// TIA Portal V20 export
// export: Created 2026-10-20T12:44:30.4346877Z, ExportSetting WithDefaults, DisplayName Totally Integrated Automation Portal, DisplayVersion V20 Update 6, DisplayName TIA Portal Openness, DisplayVersion V20 Update 6, DisplayName TIA Portal Version Control Interface, DisplayVersion V20 Update 6, DisplayName SINAMICS Startdrive Advanced, DisplayVersion V20 SP1, DisplayName SINAMICS Startdrive G130, G150, S120, S150, SINAMICS MV, G220, S200, S210, DisplayVersion V20 SP1, DisplayName SINAMICS Startdrive G110M, G120, G120C, G120D, G120P, G115D, DisplayVersion V20 SP1, DisplayName STEP 7 Professional, DisplayVersion V20 Update 6, DisplayName STEP 7 Safety, DisplayVersion V20 Update 2, DisplayName WinCC Basic/Comfort/Advanced, DisplayVersion V20 Update 6, DisplayName WinCC Unified, DisplayVersion V20 Update 6
FUNCTION "Local_Mode_FC" : Bool   // FC67, SCL
{ S7_Optimized_Access := 'TRUE' }
VERSION : 0.1
// stored: AutoNumber true, IsIECCheckEnabled false, SetENOAutomatically false, UDAEnableTagReadback false
   VAR_INPUT
      HMI_Box_Connected : Int;
      Rem_Loc_Keys : Array[1..5] of "Level_Keys_UDT";
   END_VAR
   VAR_TEMP
      System : UInt;
      Level : UInt;
   END_VAR
BEGIN
   #System := #HMI_Box_Connected / 10;
   #Level := #HMI_Box_Connected MOD 10;
   IF #System <> 0 AND #Level <> 0 THEN
       #Local_Mode_FC := #Rem_Loc_Keys[#System].Level[#Level];
   ELSE
       #Local_Mode_FC := FALSE;
   END_IF;
END_FUNCTION
